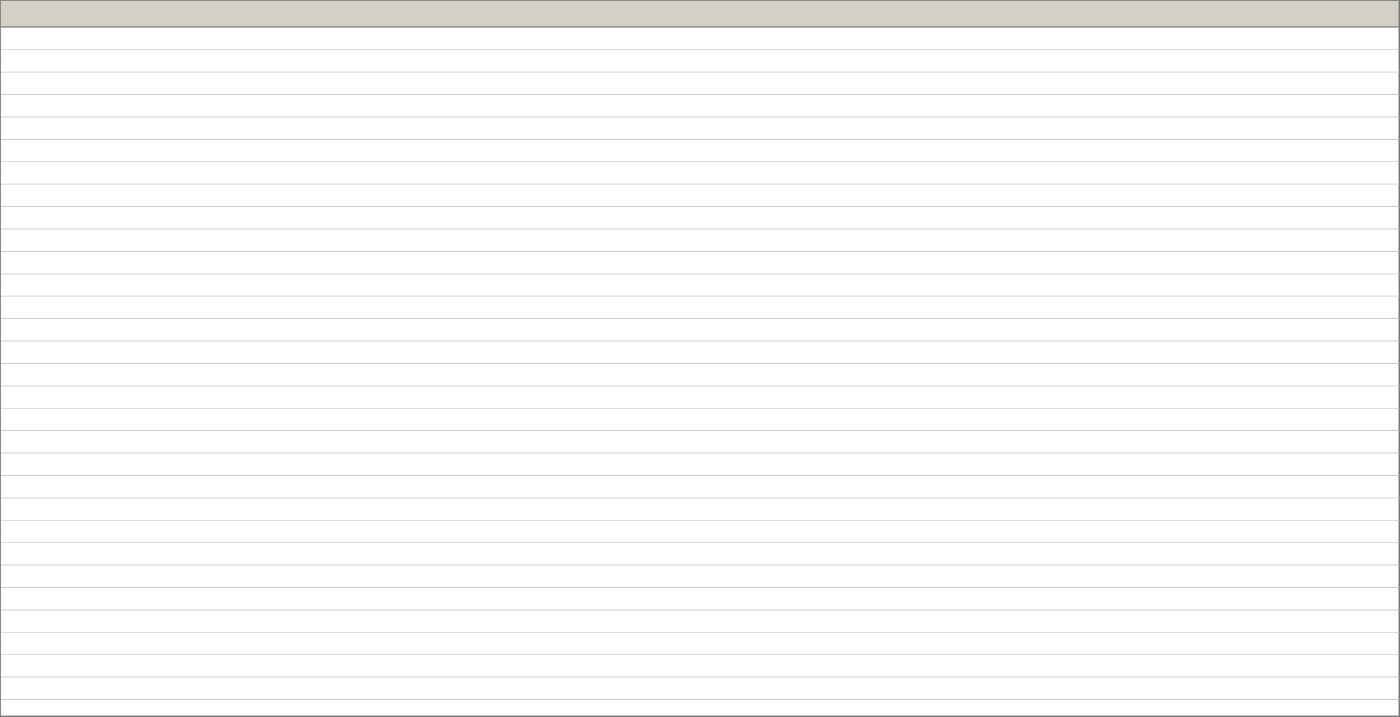
VISUALIZATION vis_Error_Act  // 1560x800
    Table (0,0 1560x800), data array: Buffer_Act_Message
        p3854506369: Buffer_Act_Message[INDEX].sDateTime
        p1892666644: Buffer_Act_Message[INDEX].sErrID
        p338671338: Buffer_Act_Message[INDEX].sLevel
        p2170511999: Buffer_Act_Message[INDEX].sModuleDescription
        p3723444502: Buffer_Act_Message[INDEX].sErrorMessage
        p4092479075: Module Description
        p2237128397: Error Message
END_VISUALIZATION

(* stored: Version 1.1.0.1, ProductVersion 3.1.4024.13
   Visu vis_Error_Act: Id {1763c5ea-f904-4a08-84ab-2f824ccd53cf} *)
